(* IEC 61131-3 sources: LASAL/Network/HW_Network, 1 file *)

(* ---- ONE_HW_Network_Table.st ---- *)
#define OBJECTS_CONFIG

//Define part of class SdiasBase
//Address to access the Dataobject list via SPI SDO Read
#define SDIAS_SPI_DATA_OBJECT_LIST_PAGE_ADDRESS 16#FFFF
#define SDIAS_SPI_DATA_OBJECT_LIST_PAGE_OFFSET 16#00
#define SDIAS_SPI_DATA_OBJECT_LIST_IDENTIFIER 16#12345678

//Defines the number of optional list elements in the SPI List

#define SDIAS_SPI_NUMBER_OF_OPTIONAL_ELEMENTS 7

//#pragma message("EisMic 27.06.2014 14:44 \ Noch schauen ob ichs besser machen kann")
#define SDIAS_SPI_HEADER_BEFORE_OPTIONAL_ELEMENTS 16#18
#define SDIAS_SPI_HARDWARE_VERSION_OFFSET 16#C
#define SDIAS_SPI_VENDOR_ID_OFFSET 16#0

//SPI List IDs
#define SDIAS_SPI_IDENTIFICATION_LIST_ID 1
#define SDIAS_SPI_FLASH_CONFIGURATION_ID 2
#define SDIAS_SPI_VENDOR_NAME_ID 3
#define SDIAS_SPI_DEVICE_NAME_ID 4
#define SDIAS_SPI_SERIAL_NUMBER_ID 5
#define SDIAS_SPI_ORDERING_NUMBER_ID 6
#define SDIAS_SPI_DOCUMENTATION_PDF_ID 7
#define SDIAS_SPI_CALIB_DATA_ID 10
#define SDIAS_SPI_PDO_INFORMATION_ID 128
#include "..\..\Class\SdiasManager\SdiasManager.h"
#include "..\..\Class\SdiasBase\SdiasBase.h"
#include "..\..\Class\HwControl\HwControl.h"
#include "..\..\Source\interfaces\lsl_st_hardwaretree.h"
#include "..\..\Source\interfaces\lsl_st_mt.h"
//Define part of class _BusInterfaceSdiasDriveMng
#define BUSIF_SDIASDRIVEMNG_OFFSET_TYPELABEL        0x0000
#define BUSIF_SDIASDRIVEMNG_PARALIST_INDEX_SET      0x2210
#define BUSIF_SDIASDRIVEMNG_PARALIST_INDEX_INFO     0x2211
#define BUSIF_SDIASDRIVEMNG_PARALIST_INDEX_SETNR    174

#define BUSIF_SDIASDRIVEMNG_MAX_SERVICEBOX          4
#define BUSIF_SDIASDRIVEMNG_SDO_RESPONSE_TIMEOUT    SDIAS_SDO_TIMEOUT * 2
#define BUSIF_SDIASDRIVEMNG_SDO_TYPELABEL_TIMEOUT   10000  //10 sec timeout to read typelabel

#define BUSIF_SDIASDRIVEMNG_SDO_SERVICE_APP_MDD100        0x4150
#define BUSIF_SDIASDRIVEMNG_SDO_SERVICE_APP_LASAL         0x4C41
#define BUSIF_SDIASDRIVEMNG_SDO_SERVICE_APP_CANOPEN       0x4453
#define BUSIF_SDIASDRIVEMNG_SDO_SERVICE_APP_CANOPEN_LASAL 0x444C

#define BUSIF_SDIASDRIVEMNG_FULL_PARADATA_SIZE   12
#define BUSIF_SDIASDRIVEMNG_CANOPEN_FOOTER_SIZE   4
#define BUSIF_SDIASDRIVEMNG_LASAL_PARADATA_SIZE   4
#include "..\..\class\_drivemngbase\drivemngbase.h"
//Define part of class _DriveAxisBase
// Device ID for the Drive Cards
#define DRIVEMNG_AXISDEVICEID_SDD_OFFSET         0
#define DRIVEMNG_AXISEVICEID_MDD_OFFSET   16#10000
#define DRIVEMNG_AXISEVICEID_SDIAS_OFFSET 16#20000
#include "..\..\Class\_DriveMngBase\SDDDefinitions.h"
//Define part of class _DriveMngBase
#ifndef _T_DRIVEMNGBASE_H
#define _T_DRIVEMNGBASE_H

// DiasDrive Constants
#DEFINE SDDMAXENTRIES   32        // maximale Anzahl an Achsen
#DEFINE SDDMAXPLACE     3         // maximale Anzahl an Achsen pro Steckplatz

// Device ID for the Drive IF Cards
#define DRIVEMNG_BUSDEVICEID_VAC011    11
#define DRIVEMNG_BUSDEVICEID_VAC012  1061
#define DRIVEMNG_BUSDEVICEID_VAC013  1075

#define DRIVEMNG_BUSDEVICEID_MDD     1071

// Device ID for the Drive Cards
#define DRIVEMNG_DRVDEVICEID_SDD_OFFSET 0

#define DRIVEMNG_DRVDEVICEID_SDD305 DRIVEMNG_DRVDEVICEID_SDD_OFFSET + 16
#define DRIVEMNG_DRVDEVICEID_SDD310 DRIVEMNG_DRVDEVICEID_SDD_OFFSET +  3
#define DRIVEMNG_DRVDEVICEID_SDD315 DRIVEMNG_DRVDEVICEID_SDD_OFFSET +  1
#define DRIVEMNG_DRVDEVICEID_SDD335 DRIVEMNG_DRVDEVICEID_SDD_OFFSET + 12

#define DRIVEMNG_DRVDEVICEID_SDD205 DRIVEMNG_DRVDEVICEID_SDD_OFFSET + 22
#define DRIVEMNG_DRVDEVICEID_SDD210 DRIVEMNG_DRVDEVICEID_SDD_OFFSET +  9
#define DRIVEMNG_DRVDEVICEID_SDD215 DRIVEMNG_DRVDEVICEID_SDD_OFFSET +  5

#define DRIVEMNG_DRVDEVICEID_SDD105 DRIVEMNG_DRVDEVICEID_SDD_OFFSET + 21
#define DRIVEMNG_DRVDEVICEID_SDD115 DRIVEMNG_DRVDEVICEID_SDD_OFFSET + 10
#define DRIVEMNG_DRVDEVICEID_SDD120 DRIVEMNG_DRVDEVICEID_SDD_OFFSET +  7

#define DRIVEMNG_DRVDEVICEID_MDD_OFFSET 16#10000

#define DRIVEMNG_DRVDEVICEID_MDD111 DRIVEMNG_DRVDEVICEID_MDD_OFFSET + 1
#define DRIVEMNG_DRVDEVICEID_MDD121 DRIVEMNG_DRVDEVICEID_MDD_OFFSET + 2

#define DRIVEMNG_DRVDEVICEID_SDIAS_OFFSET 16#20000

#define DRIVEMNG_DRVDEVICEID_DC061 DRIVEMNG_DRVDEVICEID_SDIAS_OFFSET + 16#180 // 1 = 1 Achse 80 SDIAS

#define DRIVEMNG_DRIVESCOPE_GETALL_PARAM    16#2080
#define DRIVEMNG_DRIVESCOPE_SCOPE_BIT       16#60000000
#define DRIVEMNG_DRIVESCOPE_SINDEX_RANGE    511

#endif // _T_DRIVEMNGBASE_H
//Define part of class BusInterfaceSDIASInternal
#define BUSIF_INTERNAL_MAX_NR_DO 100

// Defines for Mutex Generation
#define INTERNAL_STR_MUTEX_NAME_SEPERATOR ".."
#define INTERNAL_MUTEX_NAME_END_LENGTH 5
#define INTERNAL_MUTEX_NAME_MAX_LENGTH 32
#include "..\..\Source\BusInterface.h"
//Define part of class DM161
#define DEVICE_ID_DM161 1029
#include "..\..\Class\HwControl\watchdog.h"
#include "..\..\Source\interfaces\lsl_st_sysinfo.h"
#include "..\..\Source\interfaces\lsl_st_systrace.h"
#include <.\lsl_st_mt.h>
//Define part of class SafetyUDP
#define SAFETY_UDP_MAX_SOCKETS                6     // Max number of socket

#define SAFETY_UDP_CLT_SEND_OK                0    // Send ok
#define SAFETY_UDP_CLT_INVALID_HANDLE        -1    // Invalid handle
#define SAFETY_UDP_CLT_NOT_OPEN              -2    // Socket is not open
#define SAFETY_UDP_CLT_SEND_FAILED           -3    // Send failed
#define SAFETY_UDP_CLT_SEND_BUFFER_FULL      -4    // Send buffer is full
#define SAFETY_UDP_CLT_DATA_TO_BIG           -5    // Data to big

#define SAFETY_UDP_MAXIMUM_SEGMENT_SIZE    1452    // Maximum of user data

#define SAFETY_UDP_TIMEOUT_OPENSOCKET    (1000)    //timeout for opening socket

#define SAFETY_UDP_RECEIVE_TIMEOUT          800

#define SAFETY_UDP_TX_BUFFER_SIZE          1024
//Define part of class SafetyManager
#define LogBufferSize 1000
#include "..\..\Class\SafetyManager\SafetyManager.h"
#include "..\..\Source\interfaces\lsl_st_safetydll.h"
//Define part of class SdiasManager
#define SDIAS_SDO_MAX_LENGTH              128
#define SDIAS_SDO_RINGBUFFER_NO            64
#define SDIAS_SDO_CHANNEL_NO                3   // fixed in the VI hardware to be 3

// watchdog trigger interval (after 130ms of no trigger the SDIAS HW goes into reset again and takes at least another 10ms to be ready again)
#define SDIAS_WATCHDOG_TRIGGER_TIME        40

// time needed by sdias modules to start up after the watchdog is triggered the first time in ms
#define SDIAS_HARDWARE_STARTUP_TIME        15

// sdias manager needs 2 ticks to handle event for read task (measure sync time)
#define SDIAS_SYNC_MEASURE_TICKS            2

// after activating the PLL SyncOut it takes 3 cycles until the SDIAS sync can be injected
#define SDIAS_CYCLES_WAIT_AFTER_SYNC_ENABLE 3

// wait 1 bus cycle at start to get valid numbers in the task info
#define SDIAS_TASKINFO_READY_TICKS          1

// time to wait (in ms) until other tasks in the same or lower priority than post init have done their stuff
#define SDIAS_WAIT_TIME_IN_POST_INIT        1

#define SIZE_PER_SDIAS_CLIENT               16#0400

// for far memory accesses: 1 module can hold maximum 256 1K blocks (0-255)
#define SDIAS_1K_BLOCK_NO                       256

// far memory accesses maximum length in bytes
#define SDIAS_MAX_SIZE_FAR_MEM_ACCESS           127

#define SDIAS_OFFSET_HW_CONFIG              16#FF00
#define SDIAS_OFFSET_TASK_EVENT_IDS         16#FF10
#define SDIAS_OFFSET_FEATURE_INFO           16#FF18
#define SDIAS_OFFSET_APPLI_LED_STATES       16#FF20
#define SDIAS_OFFSET_SYNC_INJECTION_CFG     16#FF3D
#define SDIAS_OFFSET_TRIGGER_UNIT_SETUP_0   16#FF41
#define SDIAS_OFFSET_TRIGGER_UNIT_SETUP_1   16#FF45
#define SDIAS_OFFSET_TASK_START_CFG_0       16#FF60
#define SDIAS_OFFSET_TASK_CONFIG_0          16#FF86
#define SDIAS_OFFSET_TASK_CONFIG_1          16#FF96
#define SDIAS_OFFSET_TASK_INFO_1            16#FF94
#define SDIAS_OFFSET_TASK_HANDSHAKE_1       16#FF9B
#define SDIAS_OFFSET_TASK_DURATION_TIME_1   16#FF9C
#define SDIAS_OFFSET_TASK_DURATION_TIME_2   16#FFAC
#define SDIAS_OFFSET_TASK_CONFIG_2          16#FFA6

#define SDIAS_RETRIES_ALLOWED         2

// mask to get global error flag out of message counter byte of SDO responses
#define SDIAS_MASK_GLOBAL_ERROR_FLAG        16#80

// mask to get message counter out of message counter byte of SDO responses
#define SDIAS_MASK_MESSAGE_COUNTER          16#3F

#define SDIAS_EVENT_MASK_ID_SYNC_OUT0       16#10
#define SDIAS_EVENT_MASK_ID_SYNC_OUT1       16#11
#define SDIAS_EVENT_MASK_ID_SYNC_OUT2       16#12
#define SDIAS_EVENT_MASK_ID_SYNC_OUT3       16#13

#define SDIAS_MANAGER_SYNC_SYNCOUT_ID       16#85
#define SDIAS_TASK_START_EVENT_SYNCOUT_ID   16#86

#define SDIAS_PLACE_NO_MODULE_ADDED_SO_FAR  16#80000000

#define SDIAS_TRIGGER_UNIT_BYTE_SIZE        2

#define SDIAS_WAIT_TIME_FIRMWARE_HANDSHAKE  5 * 1000

// if the firmware version is below this, there might be problems with SCP111 and other modules => print warning at startup
#define SDIAS_FW_VERSION_SDO_ERROR_FIXED    16#120

// if the protocol version ist below this, Control Read/Broadcast Write Command is not supported by sdiasmanager
#define SDIAS_PROTOCOLVERSION_BROADCAST     16#120

// if the cil version ist below this, Control Read/Broadcast Write Command is not supported by OS for local SDIAS.
#define SDIAS_CILVERSION_BROADCAST         16#5001

// timeout for blocking the init during initialisation (in ms)
#define SDIAS_INIT_BLOCK_TIMEOUT            20 * 1000

#define SDIAS_MUTEX_NAME_END_LENGTH 3
#define SDIAS_MUTEX_NAME_MAX_LENGTH 32
#define SDIAS_MUTEX_STR_SEPERATOR   ".."

//#define SDIAS_RT_TIME_MEASUREMENT
#ifdef SDIAS_RT_TIME_MEASUREMENT
  #pragma message("ATTENTION: SDIAS real time measurement is active and needs additional ressources in the realtime task")
#endif

(* SDIAS data object commands  *)
#define	 SDIAS_CMD_END							  0x00			(* End command										          *)
#define	 SDIAS_CMD_ACC_MEMORY				  0x01			(* Access dpram memory								      *)
#define	 SDIAS_CMD_ACC_CONTROL				0x02			(* Access dpram control memory						  *)
#define	 SDIAS_CMD_GLOBAL						  0x03			(* SDIAS global command								      *)
#define	 SDIAS_CMD_COPY_LOCAL					0x04			(* DPRAM copy command in local dpram				*)
#define	 SDIAS_CMD_JMP_LOCAL					0x05			(* DPRAM jump command in local dpram 				*)
#define  SDIAS_CMD_ACC_MEMORY_FAR     0x07      (* SDIAS Far Memory Access                  *)

(* SDIAS defines for data object handling *)
// Write data oject list
#define	 SDIAS_DOL_WRITE_USAGE_DOL_EMPTY	  0x20			(* Usage of empty write dol list (wachtdog trigger + end command)   *)
#define	 SDIAS_DOL_WRITE_USAGE_DTA_EMPTY	  0x03			(* Usage of empty write dol data (DO ctrl of 2x copy command for task information + DO ctrl of watchdog trigger      *)
#define	 SDIAS_DOL_WRITE_OFFSET_END_CMD			0x10			(* One data object in list - offset = 1 DO size = 0x10						  *)
#define	 SDIAS_DOL_WRITE_OFFSET_FIRST_DTA		0x02			(* Offset of first data byte of second copy command = 2 (DO ctrl)   *)
#define	 SDIAS_DOL_WRITE_OFFSET_LAST_DTA		0x02			(* Offset of last data byte of second copy command = 2 (DO ctrl )   *)

// Read data oject list
#define	 SDIAS_DOL_READ_USAGE_DOL_EMPTY	    0x30			(* Usage of empty read dol list (2x task info copy command + end command)   *)
#define	 SDIAS_DOL_READ_USAGE_DTA_EMPTY	    0x0D			(* Usage of empty write dol data (DO ctrl of 2x copy command for task information + DO ctrl of watchdog trigger      *)
#define	 SDIAS_DOL_READ_OFFSET_END_CMD			0x20			(* One data object in list - offset = 1 DO size = 0x10						          *)
#define	 SDIAS_DOL_READ_OFFSET_FIRST_DTA		0x07			(* Offset of first data byte of second copy command = 7 = DO state          *)
#define	 SDIAS_DOL_READ_OFFSET_LAST_DTA		  0x0C			(* Offset of last data byte of second copy command = 12 (last byte of task information)       *)

//Versionsnumber where SDIAS SPI Read Accesses are available
#define  SDIAS_SDO_SPI_FIRMWARE_VERSION_AVAILABLE 16#0120

//error info mask
#define  SDIAS_ERROR_INFO_MASK    2#1000011000011111

// Broadcast DO Info
#define SDIAS_OFFSET_CLIENT_CTRLTIMESTAMP   16#0190
#define SDIAS_NR_TIMEBROADCAST_DOS 2
#define SDIAS_TIMEBROADCAST_SUBCMD 16#B0
#include "..\..\Source\interfaces\lsl_st_pll.h"
//Define part of class SdiasPLC
#define SDIASM_OBJECT_PATH            16#88000002   // Object Path for VSDIASmanager Length = 2 (First 2byte), Domain = 0 (3rd byte), Escape Sequence SDIAS (4th byte)
//Define part of class SR022
#define DEVICE_ID_SR022             1083        //DeviceID of SR022

#define SR022_ADDR_CYC_WRITE        16#00       //Address for TPDO
#define SR022_ADDR_CYC_READ         16#08       //Address for RPDO

#define SR022_ADDR_CFG_FIRMWARE     16#200      //Address-Offset to the Configuration of the Firmware
#define SR022_ADDR_STATE_FIRMWARE   16#280      //Address-Offset to the Status of the Firmware
#define SR022_ADDR_READ_SDO         16#0C       //Address-Offset read sdo data
#define SR022_ADDR_I2T_THRESHOLD    16#18       //Address-Offset to I²T Threshold
#define SR022_ADDR_DC_SEQUENCER     16#20       //Address-Offset to sequencer SR022

#define SR022_INVALID_VALUE         16#80000010$DINT

#define SR022_NOENCODER             0
#define SR022_TTL_MODE              1
#define SR022_RS422_MODE            2

//Define for the H-Bridge
//-----------------------------------------------------------
#define SR022_GATE_A_LOW		          2#0100000000000000    //Bit-Configuration for Enable GateA Low-Switch
#define SR022_GATE_A_HIGH		          2#0001000000000000    //Bit-Configuration for Enable GateA High-Switch
#define SR022_GATE_B_LOW		          2#1000000000000000    //Bit-Configuration for Enable GateB Low-Switch
#define SR022_GATE_B_HIGH		          2#0010000000000000    //Bit-Configuration for Enable GateB High-Switch

#define SR022_MASK_CONTROL	          16#0FFF     //Mask for Output Sequence Bits
#define SR022_MASK_TIME		            16#F000     //Mask for TimeValue

#define SR022_T_SWITCH                41      //Delay Time for Switch
#define SR022_DEFAULT_SEQ_INIT        1       //Initilization for Sequencer => After 1 FPGA-Cycle switch to next Sequency

#define SR022_FPGA_FREQ_MHZ           50    //Frequency of FPGA

#define SR022_SDO_RESPONSE_TIMEOUT  SDIAS_SDO_TIMEOUT * 2     //SDO-Response Timeout

//#define SR022_I2T_THRESHOLD          16000000   //Maximal allowed I²T Value in mA²s ==> 16 A²s
//#pragma message ("TarPet: dieser Wert wurde vorest empirisch ermittelt und sollte noch genau bestimmt werden");
#define SR022_I2T_THRESHOLD          78000   //Maximal allowed I²T Value in mA²s ==> 16 A²s

#define SR022_SPEED_SCALING          10000      //Scaling of the Server Speed (0.00% to 100.00%)
#define SR022_MINPULSE_SCALING       1000       //Scaling of the Server MinPulse (0.0% to 100.0%)
//Define part of class ST011
#define DEVICE_ID_ST011 1052
#define ST011_MINIMAL_PULSEWIDTH 16#003C

#define ST011_ADDR_PDO_WRITE    16#001F
#define ST011_ADDR_SDO_WRITE_1  16#0025
#define ST011_ADDR_PDO_READ     16#0037
#define ST011_ADDR_SDO_WRITE_2  16#0042

#define ST011_FPGAVersion_PulsCntCorrect 16#12

// in MHz
#define ST011_FREQUENCY_MHZ 125

// in Hz
#define ST011_FREQUENCY_HZ (ST011_FREQUENCY_MHZ * 1000000)

#define ST011_SDO_RESPONSE_TIMEOUT  SDIAS_SDO_TIMEOUT * 2
//Define part of class ST151Base
#define DEVICE_ID_ST151                                                    1086

#define ST151_ADDR_PDO_WRITE                                            16#0000
#define ST151_ADDR_PDO_READ                                             16#0038
#define ST151_ADDR_SDO_1                                                16#0008
#define ST151_ADDR_SDO_2           (ST151_ADDR_SDO_1+sizeof(t_s_ConfigModule1))
#define ST151_ADDR_SDO_3                                (ST151_ADDR_PDO_READ+6)  //only read sdo!!!
#define ST151_ADDR_SDO_4           (ST151_ADDR_SDO_3+sizeof(t_s_ConfigModule3))
#define ST151_ADDR_SDO_5           (ST151_ADDR_SDO_4+sizeof(t_s_ConfigModule4))
#define ST151_ADDR_SDO_6           (ST151_ADDR_SDO_5+sizeof(t_s_ConfigModule5))

#define ST151_OSZI_ADDR_WRITE                                           16#0800
#define ST151_OSZI_ADDR_READ                                            16#0808
#define ST151_OSZI_ADDR_DATA                                            16#0820
#define ST151_OSZI_READPOINTER_OFFSET                                   16#0020
#define ST151_OSZI_ONE_PDOSIZE                                              126
#define ST151_OSZI_VALUES_DATA             (ST151_OSZI_ONE_PDOSIZE/sizeof(UINT))
#define ST151_OSZI_BUFFER_SIZE                                             1024
#define ST151_OSZI_MAX_SAMPLES             (ST151_OSZI_BUFFER_SIZE/sizeof(UINT))
#define ST151_OSZI_MAX_PDOREAD   ((ST151_OSZI_BUFFER_SIZE/ST151_OSZI_ONE_PDOSIZE)+1)

// in MHz
#define ST151_FREQUENCY_MHZ                             125
// in Hz
#define ST151_FREQUENCY_HZ   (ST151_FREQUENCY_MHZ * 1000000)

#define ST151_SDO_RESPONSE_TIMEOUT   (SDIAS_SDO_TIMEOUT * 2)
#define ST151_SDO_MAX_RETRYS                              3

#define ST151_MAXFREQUENCY_OUT                   2_000_000 // 2Mhz/64 max frequency of module output
#define ST151_MAXSTEPPING_MODES                          6
#define ST151_FREQLIMITS_TABLESIZE      (ST151_MAXSTEPPING_MODES*sizeof(UDINT)*2)

#define ST151_MAX_ALLOWED_PERCENT                      100 // maximum value for percent value
#define ST151_BLANKING_TIME                             10 // minimum on time of pwm (*20ns)

#define ST151_CYCLICREFRESHDATA_TIME                   200 // time to refresh asynchrone values
#define ST151_INVALID_VALUE                   16#8000_0010 // invalid value for server
#define ST151_AUTOSET_FREQUENCYLIMIT          16#0000_0000 // value for autoset limit
#define ST151_DEACTIVATE_FREQUENCYLIMIT       16#FFFF_FFFF // value for deactivate limit

#define ST151_MAX_ALLOWED_CURRENT                     5000 // max allowed current (5A) in mA, from h-bridge according to hw-documentation
#define ST151_MAX_ALLOWED_CHOPPEROFFTIME              2500 // max allowed chopper off time in 20ns steps
#define ST151_MIN_ALLOWED_CHOPPEROFFTIME              1500 // min allowed chopper off time in 20ns steps
#define ST151_STALL_CURRENT_LIMIT                     1000 // calculation for stall current in permille
#define ST151_CURRENTOFFSETADJUST_MAX                  250 // maximum current offset adjust in mA
#define ST151_CURRENTOFFSETADJUST_MIN                 -250 // minimum current offset adjust in mA

//pll settings
#define ST151_SYNC_OUT_ID                             16#03
#define ST151_PLL_OFFSET                             16#140
#define ST151_PLL_CONTROL               (ST151_PLL_OFFSET+8)

#define ST151_ERROR_BITMASK_STATE_WORD               0x013E
#define ST151_ERROR_BITMASK_EXTENDED_STATE_WORD      0xFF3E
//Define part of class VaranManager
#define SIZE_PAYLOAD_FRAME_HEADER_DO      16#38  // Const because datasize is in the Payload DOs
#define SIZE_PAYLOAD_IRQ_FRAME_HEADER_DO  16#40  // Const because datasize is in the Payload DOs

#define VM_MAX_POST_INIT_MODULES  1000

#define VM_OBJECT_PATH            16#81000002   // Object Path for Varanmanager Length = 2 (First 2byte), Domain = 0 (3rd byte), Escape Sequence Varan (4th byte)
#include "..\..\Class\VaranManager\VaranManager.h"
#include "..\..\Source\interfaces\lsl_st_kernel.h"

FUNCTION GLOBAL TAB ONE_HW_Network
-1$UINT, 0$UINT,
0$UINT, 0$UINT,

39$UDINT,
TO_UDINT(1048633017), "_BusInterfaceSdiasDriveMng", 1$UINT, 10$UINT, 4$UINT,
TO_UDINT(529317953), "_CanLib", 1$UINT, 10$UINT, 2$UINT,
TO_UDINT(912370472), "_DriveAxis", 1$UINT, 63$UINT, 4$UINT,
TO_UDINT(4124502522), "_DriveAxisBase", 1$UINT, 72$UINT, 0$UINT,
TO_UDINT(833307860), "_DriveAxisSet", 1$UINT, 20$UINT, 4$UINT,
TO_UDINT(1470062879), "_DriveMng_DC062", 1$UINT, 16$UINT, 4$UINT,
TO_UDINT(496739206), "_DriveMngBase", 1$UINT, 41$UINT, 0$UINT,
TO_UDINT(4078275645), "_SerLib", 1$UINT, 34$UINT, 2$UINT,
TO_UDINT(2897291062), "ASCII_BIN", 1$UINT, 21$UINT, 1$UINT,
TO_UDINT(3882880897), "BusInterfaceSDIASInternal", 2$UINT, 0$UINT, 0$UINT,
TO_UDINT(658879389), "CP112_IOs", 1$UINT, 0$UINT, 1$UINT,
TO_UDINT(794617671), "CriticalSection", 0$UINT, 4$UINT, 2$UINT,
TO_UDINT(4282685340), "DM161", 1$UINT, 12$UINT, 1$UINT,
TO_UDINT(3238133653), "Hub_Base", 1$UINT, 21$UINT, 0$UINT,
TO_UDINT(1770276445), "Hub_Base_Root", 2$UINT, 11$UINT, 1$UINT,
TO_UDINT(2471641665), "HwControl", 5$UINT, 2$UINT, 1$UINT,
TO_UDINT(1193052171), "HwControlBase", 1$UINT, 10$UINT, 0$UINT,
TO_UDINT(4260294091), "HWRtPostScan", 1$UINT, 0$UINT, 1$UINT,
TO_UDINT(2225119864), "MerkerEx", 1$UINT, 22$UINT, 21$UINT,
TO_UDINT(933570811), "RAMex", 1$UINT, 17$UINT, 4$UINT,
TO_UDINT(1799751072), "SafetyManager", 2$UINT, 11$UINT, 1$UINT,
TO_UDINT(3727715967), "SafetyUDP", 1$UINT, 2$UINT, 0$UINT,
TO_UDINT(3175101883), "SdiasBase", 1$UINT, 58$UINT, 0$UINT,
TO_UDINT(4173303375), "SdiasHubBase", 1$UINT, 10$UINT, 1$UINT,
TO_UDINT(2118381352), "SdiasManager", 1$UINT, 92$UINT, 1$UINT,
TO_UDINT(1159122596), "SdiasPLC", 2$UINT, 0$UINT, 1$UINT,
TO_UDINT(2317024038), "SetCurrent", 0$UINT, 0$UINT, 1$UINT,
TO_UDINT(3646514510), "SR022", 1$UINT, 2$UINT, 1$UINT,
TO_UDINT(1310079211), "ST011", 1$UINT, 11$UINT, 1$UINT,
TO_UDINT(733517784), "ST151", 1$UINT, 2$UINT, 2$UINT,
TO_UDINT(1691609973), "ST151_IntVisu", 1$UINT, 0$UINT, 2$UINT,
TO_UDINT(1832775974), "ST151Base", 1$UINT, 2$UINT, 0$UINT,
TO_UDINT(1850111279), "String", 1$UINT, 10$UINT, 17$UINT,
TO_UDINT(2898603620), "StringInternal", 1$UINT, 82$UINT, 0$UINT,
TO_UDINT(2940693151), "VaranManager", 3$UINT, 1$UINT, 0$UINT,
TO_UDINT(1989862026), "VaranManager_1", 2$UINT, 1$UINT, 1$UINT,
TO_UDINT(4035182347), "VaranManager_Base", 1$UINT, 24$UINT, 0$UINT,
TO_UDINT(3232495061), "VirtualBaseInit", 1$UINT, 3$UINT, 0$UINT,
TO_UDINT(819479645), "XXXBase_IOs", 1$UINT, 0$UINT, 0$UINT,

1$UINT, TO_UDINT(1755887647), "_DRIVEMNG_DC0621\BUSINTERFACESDIASDRIVEMNG",
1$UINT, TO_UDINT(3678180828), "_DRIVEMNG_DC0622\BUSINTERFACESDIASDRIVEMNG",
1$UINT, TO_UDINT(3048246941), "_DRIVEMNG_DC0623\BUSINTERFACESDIASDRIVEMNG",
1$UINT, TO_UDINT(1734723611), "_DRIVEMNG_DC0624\BUSINTERFACESDIASDRIVEMNG",

1$UINT, TO_UDINT(3194356815), "CP112_IOS1\_BASE\_CANLIB1",
1$UINT, TO_UDINT(661607925), "CP112_IOS1\_BASE\_CANLIB2",

_NO_ATTR, TO_UDINT(3059689190), "_DRIVEAXIS1",
_NO_ATTR, TO_UDINT(794195804), "_DRIVEAXIS2",
_NO_ATTR, TO_UDINT(1481721802), "_DRIVEAXIS3",
_NO_ATTR, TO_UDINT(3325416041), "_DRIVEAXIS4",

1$UINT, TO_UDINT(4275951967), "_DRIVEAXIS1\SDDAXSET1",
1$UINT, TO_UDINT(1732231006), "_DRIVEAXIS2\SDDAXSET1",
1$UINT, TO_UDINT(2796642462), "_DRIVEAXIS3\SDDAXSET1",
1$UINT, TO_UDINT(2408215837), "_DRIVEAXIS4\SDDAXSET1",

_NO_ATTR, TO_UDINT(243498275), "_DRIVEMNG_DC0621",
_NO_ATTR, TO_UDINT(2542415001), "_DRIVEMNG_DC0622",
_NO_ATTR, TO_UDINT(3767344143), "_DRIVEMNG_DC0623",
_NO_ATTR, TO_UDINT(2129234348), "_DRIVEMNG_DC0624",

1$UINT, TO_UDINT(3879313428), "CP112_IOS1\_BASE\_SERLIB1",
1$UINT, TO_UDINT(2117136814), "CP112_IOS1\_BASE\_SERLIB2",

1$UINT, TO_UDINT(3603645853), "VARANMANAGER_11\_BASE\ASCII_BIN1",

_NO_ATTR, TO_UDINT(222643709), "CP112_IOS1",

1$UINT, TO_UDINT(2972590922), "HWCONTROL1\SAFETYMANAGER\UDPRECEIVEDATA",
1$UINT, TO_UDINT(1868223583), "HWCONTROL1\SAFETYMANAGER\UDPSENDDATA",

_NO_ATTR, TO_UDINT(2056942671), "DM1611",

1$UINT, TO_UDINT(1776428101), "VARANMANAGER_11\HUB_BASE_ROOT0",

_NO_ATTR, TO_UDINT(2190789875), "HWCONTROL1",

1$UINT, TO_UDINT(1673205898), "HWCONTROL1\HWRTPOSTSCAN",

1$UINT, TO_UDINT(1089285877), "DM1611\_BASE\SERIALNOSTR\MERKEREX0",
1$UINT, TO_UDINT(566457232), "SR0221\_BASE\SERIALNOSTR\MERKEREX0",
1$UINT, TO_UDINT(3227848145), "ST0111\_BASE\SERIALNOSTR\MERKEREX0",
1$UINT, TO_UDINT(921637672), "ST1511\_BASE\_BASE\SERIALNOSTR\MERKEREX0",
1$UINT, TO_UDINT(3174837553), "ST1512\_BASE\_BASE\SERIALNOSTR\MERKEREX0",
1$UINT, TO_UDINT(3868254288), "_DRIVEAXIS1\MERKEREX2",
1$UINT, TO_UDINT(2138211921), "_DRIVEAXIS2\MERKEREX2",
1$UINT, TO_UDINT(3204209041), "_DRIVEAXIS3\MERKEREX2",
1$UINT, TO_UDINT(2546420754), "_DRIVEAXIS4\MERKEREX2",
1$UINT, TO_UDINT(1361534785), "_DRIVEMNG_DC0621\BUSINTERFACESDIASDRIVEMNG\_BASE\SERIALNOSTR\MERKEREX0",
1$UINT, TO_UDINT(570430050), "_DRIVEMNG_DC0621\FWDATESTRING\MERKEREX0",
1$UINT, TO_UDINT(1339808896), "_DRIVEMNG_DC0621\FWNUMSTRING\MERKEREX0",
1$UINT, TO_UDINT(925076081), "_DRIVEMNG_DC0622\BUSINTERFACESDIASDRIVEMNG\_BASE\SERIALNOSTR\MERKEREX0",
1$UINT, TO_UDINT(2048834378), "_DRIVEMNG_DC0622\FWDATESTRING\MERKEREX0",
1$UINT, TO_UDINT(960423357), "_DRIVEMNG_DC0622\FWNUMSTRING\MERKEREX0",
1$UINT, TO_UDINT(354433377), "_DRIVEMNG_DC0623\BUSINTERFACESDIASDRIVEMNG\_BASE\SERIALNOSTR\MERKEREX0",
1$UINT, TO_UDINT(4215004781), "_DRIVEMNG_DC0623\FWDATESTRING\MERKEREX0",
1$UINT, TO_UDINT(2722959209), "_DRIVEMNG_DC0623\FWNUMSTRING\MERKEREX0",
1$UINT, TO_UDINT(4213841937), "_DRIVEMNG_DC0624\BUSINTERFACESDIASDRIVEMNG\_BASE\SERIALNOSTR\MERKEREX0",
1$UINT, TO_UDINT(3391351066), "_DRIVEMNG_DC0624\FWDATESTRING\MERKEREX0",
1$UINT, TO_UDINT(3572799431), "_DRIVEMNG_DC0624\FWNUMSTRING\MERKEREX0",

1$UINT, TO_UDINT(3414815221), "_DRIVEAXIS1\RAMEX2",
1$UINT, TO_UDINT(1158084118), "_DRIVEAXIS2\RAMEX2",
1$UINT, TO_UDINT(2309813896), "_DRIVEAXIS3\RAMEX2",
1$UINT, TO_UDINT(2204762001), "_DRIVEAXIS4\RAMEX2",

1$UINT, TO_UDINT(1778590035), "HWCONTROL1\SAFETYMANAGER",

1$UINT, TO_UDINT(1007630054), "SDIASPLC1\SDIASHUBBASE1",

1$UINT, TO_UDINT(4015996540), "SDIASPLC1\SDIASMANAGER1",

_NO_ATTR, TO_UDINT(1378000520), "SDIASPLC1",

_NO_ATTR, TO_UDINT(1364947121), "SETCURRENT1",

_NO_ATTR, TO_UDINT(308402757), "SR0221",

_NO_ATTR, TO_UDINT(3024798335), "ST0111",

_NO_ATTR, TO_UDINT(201264582), "ST1511",
_NO_ATTR, TO_UDINT(2465619068), "ST1512",

1$UINT, TO_UDINT(869501406), "ST1511\ST151_INTVISU1",
1$UINT, TO_UDINT(437992748), "ST1512\ST151_INTVISU1",

1$UINT, TO_UDINT(2011818843), "DM1611\_BASE\SERIALNOSTR",
1$UINT, TO_UDINT(3834696548), "SR0221\_BASE\SERIALNOSTR",
1$UINT, TO_UDINT(3723324983), "ST0111\_BASE\SERIALNOSTR",
1$UINT, TO_UDINT(3070230801), "ST1511\_BASE\_BASE\SERIALNOSTR",
1$UINT, TO_UDINT(2196617026), "ST1512\_BASE\_BASE\SERIALNOSTR",
1$UINT, TO_UDINT(189353776), "_DRIVEMNG_DC0621\BUSINTERFACESDIASDRIVEMNG\_BASE\SERIALNOSTR",
1$UINT, TO_UDINT(275191107), "_DRIVEMNG_DC0621\FWDATESTRING",
1$UINT, TO_UDINT(1236665617), "_DRIVEMNG_DC0621\FWNUMSTRING",
1$UINT, TO_UDINT(880947621), "_DRIVEMNG_DC0622\BUSINTERFACESDIASDRIVEMNG\_BASE\SERIALNOSTR",
1$UINT, TO_UDINT(1812344984), "_DRIVEMNG_DC0622\FWDATESTRING",
1$UINT, TO_UDINT(4101794271), "_DRIVEMNG_DC0622\FWNUMSTRING",
1$UINT, TO_UDINT(2534676969), "_DRIVEMNG_DC0623\BUSINTERFACESDIASDRIVEMNG\_BASE\SERIALNOSTR",
1$UINT, TO_UDINT(4043952622), "_DRIVEMNG_DC0623\FWDATESTRING",
1$UINT, TO_UDINT(703246426), "_DRIVEMNG_DC0623\FWNUMSTRING",
1$UINT, TO_UDINT(1259654287), "_DRIVEMNG_DC0624\BUSINTERFACESDIASDRIVEMNG\_BASE\SERIALNOSTR",
1$UINT, TO_UDINT(2495904558), "_DRIVEMNG_DC0624\FWDATESTRING",
1$UINT, TO_UDINT(1419359746), "_DRIVEMNG_DC0624\FWNUMSTRING",

_NO_ATTR, TO_UDINT(2395414379), "VARANMANAGER_11",

//Internal connections
0$UDINT,
64$UDINT,
TO_UDINT(0), "SerialNoStr", TO_UDINT(69),
TO_UDINT(1), "SerialNoStr", TO_UDINT(72),
TO_UDINT(2), "SerialNoStr", TO_UDINT(75),
TO_UDINT(3), "SerialNoStr", TO_UDINT(78),
TO_UDINT(6), "SDDAxSet1", TO_UDINT(10),
TO_UDINT(6), "MerkerEx2", TO_UDINT(33),
TO_UDINT(6), "RAMex2", TO_UDINT(49),
TO_UDINT(7), "SDDAxSet1", TO_UDINT(11),
TO_UDINT(7), "MerkerEx2", TO_UDINT(34),
TO_UDINT(7), "RAMex2", TO_UDINT(50),
TO_UDINT(8), "SDDAxSet1", TO_UDINT(12),
TO_UDINT(8), "MerkerEx2", TO_UDINT(35),
TO_UDINT(8), "RAMex2", TO_UDINT(51),
TO_UDINT(9), "SDDAxSet1", TO_UDINT(13),
TO_UDINT(9), "MerkerEx2", TO_UDINT(36),
TO_UDINT(9), "RAMex2", TO_UDINT(52),
TO_UDINT(14), "FWDateString", TO_UDINT(70),
TO_UDINT(14), "FWNumSTring", TO_UDINT(71),
TO_UDINT(14), "BusInterfaceSdiasDriveMng", TO_UDINT(0),
TO_UDINT(15), "FWDateString", TO_UDINT(73),
TO_UDINT(15), "FWNumSTring", TO_UDINT(74),
TO_UDINT(15), "BusInterfaceSdiasDriveMng", TO_UDINT(1),
TO_UDINT(16), "FWDateString", TO_UDINT(76),
TO_UDINT(16), "FWNumSTring", TO_UDINT(77),
TO_UDINT(16), "BusInterfaceSdiasDriveMng", TO_UDINT(2),
TO_UDINT(17), "FWDateString", TO_UDINT(79),
TO_UDINT(17), "FWNumSTring", TO_UDINT(80),
TO_UDINT(17), "BusInterfaceSdiasDriveMng", TO_UDINT(3),
TO_UDINT(21), "_SerLib1", TO_UDINT(18),
TO_UDINT(21), "_SerLib2", TO_UDINT(19),
TO_UDINT(21), "_CanLib1", TO_UDINT(4),
TO_UDINT(21), "_CanLib2", TO_UDINT(5),
TO_UDINT(24), "SerialNoStr", TO_UDINT(64),
TO_UDINT(26), "SafetyManager", TO_UDINT(53),
TO_UDINT(26), "HWRtPostScan", TO_UDINT(27),
TO_UDINT(53), "UdpSendData", TO_UDINT(23),
TO_UDINT(53), "UdpReceiveData", TO_UDINT(22),
TO_UDINT(56), "SdiasManager1", TO_UDINT(55),
TO_UDINT(56), "SdiasHubBase1", TO_UDINT(54),
TO_UDINT(58), "SerialNoStr", TO_UDINT(65),
TO_UDINT(59), "SerialNoStr", TO_UDINT(66),
TO_UDINT(60), "SerialNoStr", TO_UDINT(67),
TO_UDINT(60), "ST151_IntVisu1", TO_UDINT(62),
TO_UDINT(61), "SerialNoStr", TO_UDINT(68),
TO_UDINT(61), "ST151_IntVisu1", TO_UDINT(63),
TO_UDINT(64), "MerkerEx0", TO_UDINT(28),
TO_UDINT(65), "MerkerEx0", TO_UDINT(29),
TO_UDINT(66), "MerkerEx0", TO_UDINT(30),
TO_UDINT(67), "MerkerEx0", TO_UDINT(31),
TO_UDINT(68), "MerkerEx0", TO_UDINT(32),
TO_UDINT(69), "MerkerEx0", TO_UDINT(37),
TO_UDINT(70), "MerkerEx0", TO_UDINT(38),
TO_UDINT(71), "MerkerEx0", TO_UDINT(39),
TO_UDINT(72), "MerkerEx0", TO_UDINT(40),
TO_UDINT(73), "MerkerEx0", TO_UDINT(41),
TO_UDINT(74), "MerkerEx0", TO_UDINT(42),
TO_UDINT(75), "MerkerEx0", TO_UDINT(43),
TO_UDINT(76), "MerkerEx0", TO_UDINT(44),
TO_UDINT(77), "MerkerEx0", TO_UDINT(45),
TO_UDINT(78), "MerkerEx0", TO_UDINT(46),
TO_UDINT(79), "MerkerEx0", TO_UDINT(47),
TO_UDINT(80), "MerkerEx0", TO_UDINT(48),
TO_UDINT(81), "ASCII_BIN1", TO_UDINT(20),
TO_UDINT(81), "Hub_Base_Root0", TO_UDINT(25),
0$UDINT,
69$UDINT,
TO_UDINT(6), "DriveMng", TO_UDINT(14), "CmdState",
TO_UDINT(6), "DriveAxisSet", TO_UDINT(10), "Server0",
TO_UDINT(7), "DriveMng", TO_UDINT(15), "CmdState",
TO_UDINT(7), "DriveAxisSet", TO_UDINT(11), "Server0",
TO_UDINT(8), "DriveMng", TO_UDINT(16), "CmdState",
TO_UDINT(8), "DriveAxisSet", TO_UDINT(12), "Server0",
TO_UDINT(9), "DriveMng", TO_UDINT(17), "CmdState",
TO_UDINT(9), "DriveAxisSet", TO_UDINT(13), "Server0",
TO_UDINT(10), "coMerkerEx", TO_UDINT(33), "m_udLength",
TO_UDINT(10), "coRamEx", TO_UDINT(49), "m_udLength",
TO_UDINT(11), "coMerkerEx", TO_UDINT(34), "m_udLength",
TO_UDINT(11), "coRamEx", TO_UDINT(50), "m_udLength",
TO_UDINT(12), "coMerkerEx", TO_UDINT(35), "m_udLength",
TO_UDINT(12), "coRamEx", TO_UDINT(51), "m_udLength",
TO_UDINT(13), "coMerkerEx", TO_UDINT(36), "m_udLength",
TO_UDINT(13), "coRamEx", TO_UDINT(52), "m_udLength",
TO_UDINT(14), "cOnline", TO_UDINT(0), "Online",
TO_UDINT(14), "FwNumStr", TO_UDINT(71), "Data",
TO_UDINT(14), "FwDatetr", TO_UDINT(70), "Data",
TO_UDINT(14), "ToBusIF", TO_UDINT(0), "CallCommand",
TO_UDINT(14), "SdiasIn", TO_UDINT(54), "ClassSvr",
TO_UDINT(15), "cOnline", TO_UDINT(1), "Online",
TO_UDINT(15), "FwNumStr", TO_UDINT(74), "Data",
TO_UDINT(15), "FwDatetr", TO_UDINT(73), "Data",
TO_UDINT(15), "ToBusIF", TO_UDINT(1), "CallCommand",
TO_UDINT(15), "SdiasIn", TO_UDINT(54), "ClassSvr",
TO_UDINT(16), "cOnline", TO_UDINT(2), "Online",
TO_UDINT(16), "FwNumStr", TO_UDINT(77), "Data",
TO_UDINT(16), "FwDatetr", TO_UDINT(76), "Data",
TO_UDINT(16), "ToBusIF", TO_UDINT(2), "CallCommand",
TO_UDINT(16), "SdiasIn", TO_UDINT(54), "ClassSvr",
TO_UDINT(17), "cOnline", TO_UDINT(3), "Online",
TO_UDINT(17), "FwNumStr", TO_UDINT(80), "Data",
TO_UDINT(17), "FwDatetr", TO_UDINT(79), "Data",
TO_UDINT(17), "ToBusIF", TO_UDINT(3), "CallCommand",
TO_UDINT(17), "SdiasIn", TO_UDINT(54), "ClassSvr",
TO_UDINT(21), "To_HwControl", TO_UDINT(26), "Control",
TO_UDINT(24), "SdiasIn", TO_UDINT(54), "ClassSvr",
TO_UDINT(25), "VaranConnect", TO_UDINT(81), "Control",
TO_UDINT(27), "toHwControlBase", TO_UDINT(26), "Control",
TO_UDINT(53), "To_HwControl", TO_UDINT(26), "Control",
TO_UDINT(54), "ToNextSDIAS", TO_UDINT(55), "ClassState",
TO_UDINT(55), "ToBusInterface", TO_UDINT(56), "CallCommand",
TO_UDINT(56), "ToHwControl", TO_UDINT(26), "Control",
TO_UDINT(57), "Current", TO_UDINT(60), "MaxCurrent",
TO_UDINT(58), "SdiasIn", TO_UDINT(54), "ClassSvr",
TO_UDINT(59), "SdiasIn", TO_UDINT(54), "ClassSvr",
TO_UDINT(60), "SdiasIn", TO_UDINT(54), "ClassSvr",
TO_UDINT(61), "SdiasIn", TO_UDINT(54), "ClassSvr",
TO_UDINT(62), "toST151Base", TO_UDINT(60), "ClassState",
TO_UDINT(63), "toST151Base", TO_UDINT(61), "ClassState",
TO_UDINT(64), "DataBuffer", TO_UDINT(28), "m_udLength",
TO_UDINT(65), "DataBuffer", TO_UDINT(29), "m_udLength",
TO_UDINT(66), "DataBuffer", TO_UDINT(30), "m_udLength",
TO_UDINT(67), "DataBuffer", TO_UDINT(31), "m_udLength",
TO_UDINT(68), "DataBuffer", TO_UDINT(32), "m_udLength",
TO_UDINT(69), "DataBuffer", TO_UDINT(37), "m_udLength",
TO_UDINT(70), "DataBuffer", TO_UDINT(38), "m_udLength",
TO_UDINT(71), "DataBuffer", TO_UDINT(39), "m_udLength",
TO_UDINT(72), "DataBuffer", TO_UDINT(40), "m_udLength",
TO_UDINT(73), "DataBuffer", TO_UDINT(41), "m_udLength",
TO_UDINT(74), "DataBuffer", TO_UDINT(42), "m_udLength",
TO_UDINT(75), "DataBuffer", TO_UDINT(43), "m_udLength",
TO_UDINT(76), "DataBuffer", TO_UDINT(44), "m_udLength",
TO_UDINT(77), "DataBuffer", TO_UDINT(45), "m_udLength",
TO_UDINT(78), "DataBuffer", TO_UDINT(46), "m_udLength",
TO_UDINT(79), "DataBuffer", TO_UDINT(47), "m_udLength",
TO_UDINT(80), "DataBuffer", TO_UDINT(48), "m_udLength",
TO_UDINT(81), "To_HwControl", TO_UDINT(26), "Control",

//Initialization values
0$UDINT,
232$UDINT,
TO_UDINT(0), "LEDControl", TO_UDINT(0),//|HW_Network._DriveMng_DC0621\BusInterfaceSdiasDriveMng.LEDControl;
TO_UDINT(0), "Place", TO_UDINT(0),//|HW_Network._DriveMng_DC0621\BusInterfaceSdiasDriveMng.Place;
TO_UDINT(0), "Required", TO_UDINT(1),//|HW_Network._DriveMng_DC0621\BusInterfaceSdiasDriveMng.Required;
TO_UDINT(0), "TimeMultiplier", TO_UDINT(1),//|HW_Network._DriveMng_DC0621\BusInterfaceSdiasDriveMng.TimeMultiplier;
TO_UDINT(0), "SdiasID", TO_UDINT(1801),//|HW_Network._DriveMng_DC0621\BusInterfaceSdiasDriveMng.SdiasID;
TO_UDINT(1), "LEDControl", TO_UDINT(0),//|HW_Network._DriveMng_DC0622\BusInterfaceSdiasDriveMng.LEDControl;
TO_UDINT(1), "Place", TO_UDINT(1),//|HW_Network._DriveMng_DC0622\BusInterfaceSdiasDriveMng.Place;
TO_UDINT(1), "Required", TO_UDINT(1),//|HW_Network._DriveMng_DC0622\BusInterfaceSdiasDriveMng.Required;
TO_UDINT(1), "TimeMultiplier", TO_UDINT(1),//|HW_Network._DriveMng_DC0622\BusInterfaceSdiasDriveMng.TimeMultiplier;
TO_UDINT(1), "SdiasID", TO_UDINT(1801),//|HW_Network._DriveMng_DC0622\BusInterfaceSdiasDriveMng.SdiasID;
TO_UDINT(2), "LEDControl", TO_UDINT(0),//|HW_Network._DriveMng_DC0623\BusInterfaceSdiasDriveMng.LEDControl;
TO_UDINT(2), "Place", TO_UDINT(2),//|HW_Network._DriveMng_DC0623\BusInterfaceSdiasDriveMng.Place;
TO_UDINT(2), "Required", TO_UDINT(1),//|HW_Network._DriveMng_DC0623\BusInterfaceSdiasDriveMng.Required;
TO_UDINT(2), "TimeMultiplier", TO_UDINT(1),//|HW_Network._DriveMng_DC0623\BusInterfaceSdiasDriveMng.TimeMultiplier;
TO_UDINT(2), "SdiasID", TO_UDINT(1801),//|HW_Network._DriveMng_DC0623\BusInterfaceSdiasDriveMng.SdiasID;
TO_UDINT(3), "LEDControl", TO_UDINT(0),//|HW_Network._DriveMng_DC0624\BusInterfaceSdiasDriveMng.LEDControl;
TO_UDINT(3), "Place", TO_UDINT(3),//|HW_Network._DriveMng_DC0624\BusInterfaceSdiasDriveMng.Place;
TO_UDINT(3), "Required", TO_UDINT(1),//|HW_Network._DriveMng_DC0624\BusInterfaceSdiasDriveMng.Required;
TO_UDINT(3), "TimeMultiplier", TO_UDINT(1),//|HW_Network._DriveMng_DC0624\BusInterfaceSdiasDriveMng.TimeMultiplier;
TO_UDINT(3), "SdiasID", TO_UDINT(1801),//|HW_Network._DriveMng_DC0624\BusInterfaceSdiasDriveMng.SdiasID;
TO_UDINT(4), "CanBus", TO_UDINT(0),//|HW_Network._base\CP112_IOs1\_CanLib1.CanBus;
TO_UDINT(5), "CanBus", TO_UDINT(1),//|HW_Network._base\CP112_IOs1\_CanLib2.CanBus;
TO_UDINT(6), "Place", TO_UDINT(0),//|HW_Network._DriveAxis1.Place;
TO_UDINT(6), "AxisNo", TO_UDINT(1),//|HW_Network._DriveAxis1.AxisNo;
TO_UDINT(6), "AxisExtend", TO_UDINT(1),//|HW_Network._DriveAxis1.AxisExtend;
TO_UDINT(6), "ParaSaveType", TO_UDINT(1),//|HW_Network._DriveAxis1.ParaSaveType;
TO_UDINT(6), "OverwriteMotorPara", TO_UDINT(1),//|HW_Network._DriveAxis1.OverwriteMotorPara;
TO_UDINT(7), "Place", TO_UDINT(0),//|HW_Network._DriveAxis2.Place;
TO_UDINT(7), "AxisNo", TO_UDINT(1),//|HW_Network._DriveAxis2.AxisNo;
TO_UDINT(7), "AxisExtend", TO_UDINT(1),//|HW_Network._DriveAxis2.AxisExtend;
TO_UDINT(7), "ParaSaveType", TO_UDINT(1),//|HW_Network._DriveAxis2.ParaSaveType;
TO_UDINT(7), "OverwriteMotorPara", TO_UDINT(1),//|HW_Network._DriveAxis2.OverwriteMotorPara;
TO_UDINT(8), "Place", TO_UDINT(0),//|HW_Network._DriveAxis3.Place;
TO_UDINT(8), "AxisNo", TO_UDINT(1),//|HW_Network._DriveAxis3.AxisNo;
TO_UDINT(8), "AxisExtend", TO_UDINT(1),//|HW_Network._DriveAxis3.AxisExtend;
TO_UDINT(8), "ParaSaveType", TO_UDINT(1),//|HW_Network._DriveAxis3.ParaSaveType;
TO_UDINT(8), "OverwriteMotorPara", TO_UDINT(1),//|HW_Network._DriveAxis3.OverwriteMotorPara;
TO_UDINT(9), "Place", TO_UDINT(0),//|HW_Network._DriveAxis4.Place;
TO_UDINT(9), "AxisNo", TO_UDINT(1),//|HW_Network._DriveAxis4.AxisNo;
TO_UDINT(9), "AxisExtend", TO_UDINT(1),//|HW_Network._DriveAxis4.AxisExtend;
TO_UDINT(9), "ParaSaveType", TO_UDINT(1),//|HW_Network._DriveAxis4.ParaSaveType;
TO_UDINT(9), "OverwriteMotorPara", TO_UDINT(1),//|HW_Network._DriveAxis4.OverwriteMotorPara;
TO_UDINT(10), "ParaSaveType", TO_UDINT(1),//|HW_Network._DriveAxis1\SDDAxSet1.ParaSaveType;
TO_UDINT(10), "OverwriteMotorPara", TO_UDINT(1),//|HW_Network._DriveAxis1\SDDAxSet1.OverwriteMotorPara;
TO_UDINT(11), "ParaSaveType", TO_UDINT(1),//|HW_Network._DriveAxis2\SDDAxSet1.ParaSaveType;
TO_UDINT(11), "OverwriteMotorPara", TO_UDINT(1),//|HW_Network._DriveAxis2\SDDAxSet1.OverwriteMotorPara;
TO_UDINT(12), "ParaSaveType", TO_UDINT(1),//|HW_Network._DriveAxis3\SDDAxSet1.ParaSaveType;
TO_UDINT(12), "OverwriteMotorPara", TO_UDINT(1),//|HW_Network._DriveAxis3\SDDAxSet1.OverwriteMotorPara;
TO_UDINT(13), "ParaSaveType", TO_UDINT(1),//|HW_Network._DriveAxis4\SDDAxSet1.ParaSaveType;
TO_UDINT(13), "OverwriteMotorPara", TO_UDINT(1),//|HW_Network._DriveAxis4\SDDAxSet1.OverwriteMotorPara;
TO_UDINT(14), "Place", TO_UDINT(0),//|HW_Network._DriveMng_DC0621.Place;
TO_UDINT(14), "Required", TO_UDINT(1),//|HW_Network._DriveMng_DC0621.Required;
TO_UDINT(14), "TimeMultiplier", TO_UDINT(1),//|HW_Network._DriveMng_DC0621.TimeMultiplier;
TO_UDINT(15), "Place", TO_UDINT(1),//|HW_Network._DriveMng_DC0622.Place;
TO_UDINT(15), "Required", TO_UDINT(1),//|HW_Network._DriveMng_DC0622.Required;
TO_UDINT(15), "TimeMultiplier", TO_UDINT(1),//|HW_Network._DriveMng_DC0622.TimeMultiplier;
TO_UDINT(16), "Place", TO_UDINT(2),//|HW_Network._DriveMng_DC0623.Place;
TO_UDINT(16), "Required", TO_UDINT(1),//|HW_Network._DriveMng_DC0623.Required;
TO_UDINT(16), "TimeMultiplier", TO_UDINT(1),//|HW_Network._DriveMng_DC0623.TimeMultiplier;
TO_UDINT(17), "Place", TO_UDINT(3),//|HW_Network._DriveMng_DC0624.Place;
TO_UDINT(17), "Required", TO_UDINT(1),//|HW_Network._DriveMng_DC0624.Required;
TO_UDINT(17), "TimeMultiplier", TO_UDINT(1),//|HW_Network._DriveMng_DC0624.TimeMultiplier;
TO_UDINT(18), "Com", TO_UDINT(0),//|HW_Network._base\CP112_IOs1\_SerLib1.Com;
TO_UDINT(19), "Com", TO_UDINT(1),//|HW_Network._base\CP112_IOs1\_SerLib2.Com;
TO_UDINT(24), "LEDControl", TO_UDINT(0),//|HW_Network.DM1611.LEDControl;
TO_UDINT(24), "Place", TO_UDINT(4),//|HW_Network.DM1611.Place;
TO_UDINT(24), "Required", TO_UDINT(1),//|HW_Network.DM1611.Required;
TO_UDINT(25), "Splitter_Place", TO_UDINT(0),//|HW_Network.VaranManager_11\Hub_Base_Root0.Splitter_Place;
TO_UDINT(26), "UdpSafetyPort", TO_UDINT(10823),//|HW_Network.HwControl1.UdpSafetyPort;
TO_UDINT(26), "InterfaceNo", TO_UDINT(1),//|HW_Network.HwControl1.InterfaceNo;
TO_UDINT(28), "ThreadSafe", TO_UDINT(0),//|HW_Network.SerialNoStr\_base\DM1611\MerkerEx0.ThreadSafe;
TO_UDINT(29), "ThreadSafe", TO_UDINT(0),//|HW_Network.SerialNoStr\_base\SR0221\MerkerEx0.ThreadSafe;
TO_UDINT(30), "ThreadSafe", TO_UDINT(0),//|HW_Network.SerialNoStr\_base\ST0111\MerkerEx0.ThreadSafe;
TO_UDINT(31), "ThreadSafe", TO_UDINT(0),//|HW_Network.SerialNoStr\_base\_base\ST1511\MerkerEx0.ThreadSafe;
TO_UDINT(32), "ThreadSafe", TO_UDINT(0),//|HW_Network.SerialNoStr\_base\_base\ST1512\MerkerEx0.ThreadSafe;
TO_UDINT(33), "ThreadSafe", TO_UDINT(0),//|HW_Network._DriveAxis1\MerkerEx2.ThreadSafe;
TO_UDINT(34), "ThreadSafe", TO_UDINT(0),//|HW_Network._DriveAxis2\MerkerEx2.ThreadSafe;
TO_UDINT(35), "ThreadSafe", TO_UDINT(0),//|HW_Network._DriveAxis3\MerkerEx2.ThreadSafe;
TO_UDINT(36), "ThreadSafe", TO_UDINT(0),//|HW_Network._DriveAxis4\MerkerEx2.ThreadSafe;
TO_UDINT(37), "ThreadSafe", TO_UDINT(0),//|HW_Network.SerialNoStr\_base\BusInterfaceSdiasDriveMng\_DriveMng_DC0621\MerkerEx0.ThreadSafe;
TO_UDINT(38), "ThreadSafe", TO_UDINT(0),//|HW_Network.FWDateString\_DriveMng_DC0621\MerkerEx0.ThreadSafe;
TO_UDINT(39), "ThreadSafe", TO_UDINT(0),//|HW_Network.FWNumSTring\_DriveMng_DC0621\MerkerEx0.ThreadSafe;
TO_UDINT(40), "ThreadSafe", TO_UDINT(0),//|HW_Network.SerialNoStr\_base\BusInterfaceSdiasDriveMng\_DriveMng_DC0622\MerkerEx0.ThreadSafe;
TO_UDINT(41), "ThreadSafe", TO_UDINT(0),//|HW_Network.FWDateString\_DriveMng_DC0622\MerkerEx0.ThreadSafe;
TO_UDINT(42), "ThreadSafe", TO_UDINT(0),//|HW_Network.FWNumSTring\_DriveMng_DC0622\MerkerEx0.ThreadSafe;
TO_UDINT(43), "ThreadSafe", TO_UDINT(0),//|HW_Network.SerialNoStr\_base\BusInterfaceSdiasDriveMng\_DriveMng_DC0623\MerkerEx0.ThreadSafe;
TO_UDINT(44), "ThreadSafe", TO_UDINT(0),//|HW_Network.FWDateString\_DriveMng_DC0623\MerkerEx0.ThreadSafe;
TO_UDINT(45), "ThreadSafe", TO_UDINT(0),//|HW_Network.FWNumSTring\_DriveMng_DC0623\MerkerEx0.ThreadSafe;
TO_UDINT(46), "ThreadSafe", TO_UDINT(0),//|HW_Network.SerialNoStr\_base\BusInterfaceSdiasDriveMng\_DriveMng_DC0624\MerkerEx0.ThreadSafe;
TO_UDINT(47), "ThreadSafe", TO_UDINT(0),//|HW_Network.FWDateString\_DriveMng_DC0624\MerkerEx0.ThreadSafe;
TO_UDINT(48), "ThreadSafe", TO_UDINT(0),//|HW_Network.FWNumSTring\_DriveMng_DC0624\MerkerEx0.ThreadSafe;
TO_UDINT(49), "ThreadSafe", TO_UDINT(0),//|HW_Network._DriveAxis1\RAMex2.ThreadSafe;
TO_UDINT(50), "ThreadSafe", TO_UDINT(0),//|HW_Network._DriveAxis2\RAMex2.ThreadSafe;
TO_UDINT(51), "ThreadSafe", TO_UDINT(0),//|HW_Network._DriveAxis3\RAMex2.ThreadSafe;
TO_UDINT(52), "ThreadSafe", TO_UDINT(0),//|HW_Network._DriveAxis4\RAMex2.ThreadSafe;
TO_UDINT(53), "UdpSafetyPort", TO_UDINT(10823),//|HW_Network.HwControl1\SafetyManager.UdpSafetyPort;
TO_UDINT(53), "InterfaceNo", TO_UDINT(1),//|HW_Network.HwControl1\SafetyManager.InterfaceNo;
TO_UDINT(54), "SplitterPlace", TO_UDINT(0),//|HW_Network.SdiasPLC1\SdiasHubBase1.SplitterPlace;
TO_UDINT(55), "DeviceID", TO_UDINT(0),//|HW_Network.SdiasPLC1\SdiasManager1.DeviceID;
TO_UDINT(56), "CycleTime", TO_UDINT(1000),//|HW_Network.SdiasPLC1.CycleTime;
TO_UDINT(56), "IsoStartPoint", TO_UDINT(60),//|HW_Network.SdiasPLC1.IsoStartPoint;
TO_UDINT(58), "LEDControl", TO_UDINT(0),//|HW_Network.SR0221.LEDControl;
TO_UDINT(58), "MinPulse", TO_UDINT(7),//|HW_Network.SR0221.MinPulse;
TO_UDINT(58), "Place", TO_UDINT(6),//|HW_Network.SR0221.Place;
TO_UDINT(58), "Required", TO_UDINT(1),//|HW_Network.SR0221.Required;
TO_UDINT(58), "PWMPeriod", TO_UDINT(32),//|HW_Network.SR0221.PWMPeriod;
TO_UDINT(58), "I2TThreshold", TO_UDINT(100),//|HW_Network.SR0221.I2TThreshold;
TO_UDINT(58), "EncMode", TO_UDINT(1),//|HW_Network.SR0221.EncMode;
TO_UDINT(58), "EncSampling", TO_UDINT(3),//|HW_Network.SR0221.EncSampling;
TO_UDINT(58), "EncDirection", TO_UDINT(0),//|HW_Network.SR0221.EncDirection;
TO_UDINT(58), "InvertZeroPosition", TO_UDINT(0),//|HW_Network.SR0221.InvertZeroPosition;
TO_UDINT(58), "ABCountMode", TO_UDINT(0),//|HW_Network.SR0221.ABCountMode;
TO_UDINT(58), "ExtendedData", TO_UDINT(0),//|HW_Network.SR0221.ExtendedData;
TO_UDINT(59), "LEDControl", TO_UDINT(0),//|HW_Network.ST0111.LEDControl;
TO_UDINT(59), "Place", TO_UDINT(8),//|HW_Network.ST0111.Place;
TO_UDINT(59), "Required", TO_UDINT(1),//|HW_Network.ST0111.Required;
TO_UDINT(59), "UsePulseCntCorrection", TO_UDINT(1),//|HW_Network.ST0111.UsePulseCntCorrection;
TO_UDINT(59), "PulseMode", TO_UDINT(0),//|HW_Network.ST0111.PulseMode;
TO_UDINT(59), "ModeClockCounter", TO_UDINT(0),//|HW_Network.ST0111.ModeClockCounter;
TO_UDINT(59), "InvertEncoder", TO_UDINT(1),//|HW_Network.ST0111.InvertEncoder;
TO_UDINT(59), "InvertEnable", TO_UDINT(1),//|HW_Network.ST0111.InvertEnable;
TO_UDINT(59), "EncoderSampling", TO_UDINT(3),//|HW_Network.ST0111.EncoderSampling;
TO_UDINT(59), "Deathtime", TO_UDINT(60),//|HW_Network.ST0111.Deathtime;
TO_UDINT(59), "Input1Latch", TO_UDINT(0),//|HW_Network.ST0111.Input1Latch;
TO_UDINT(59), "Input2Latch", TO_UDINT(0),//|HW_Network.ST0111.Input2Latch;
TO_UDINT(59), "Input3Latch", TO_UDINT(0),//|HW_Network.ST0111.Input3Latch;
TO_UDINT(59), "ZPulseLatch", TO_UDINT(0),//|HW_Network.ST0111.ZPulseLatch;
TO_UDINT(60), "LEDControl", TO_UDINT(0),//|HW_Network.ST1511.LEDControl;
TO_UDINT(60), "CurrentIncrease", TO_UDINT(1),//|HW_Network.ST1511.CurrentIncrease;
TO_UDINT(60), "HWRampdownDeltaFrequency", TO_UDINT(40),//|HW_Network.ST1511.HWRampdownDeltaFrequency;
TO_UDINT(60), "HWRampdownDeltaTime", TO_UDINT(1),//|HW_Network.ST1511.HWRampdownDeltaTime;
TO_UDINT(60), "CurrentOffsetAdjBridge1", TO_UDINT(100),//|HW_Network.ST1511.CurrentOffsetAdjBridge1;
TO_UDINT(60), "CurrentOffsetAdjBridge2", TO_UDINT(100),//|HW_Network.ST1511.CurrentOffsetAdjBridge2;
TO_UDINT(60), "ChopperOffTime", TO_UDINT(1562),//|HW_Network.ST1511.ChopperOffTime;
TO_UDINT(60), "ChopperOnTimeMin", TO_UDINT(180),//|HW_Network.ST1511.ChopperOnTimeMin;
TO_UDINT(60), "FastDecayTime", TO_UDINT(200),//|HW_Network.ST1511.FastDecayTime;
TO_UDINT(60), "FastDecayTimeFallingStep", TO_UDINT(600),//|HW_Network.ST1511.FastDecayTimeFallingStep;
TO_UDINT(60), "EnableSteps", TO_UDINT(2#1000111),//|HW_Network.ST1511.EnableSteps;
TO_UDINT(60), "FrequLimitIncrease2to1", TO_UDINT(50000),//|HW_Network.ST1511.FrequLimitIncrease2to1;
TO_UDINT(60), "FrequLimitIncrease4to2", TO_UDINT(40000),//|HW_Network.ST1511.FrequLimitIncrease4to2;
TO_UDINT(60), "FrequLimitIncrease8to4", TO_UDINT(30000),//|HW_Network.ST1511.FrequLimitIncrease8to4;
TO_UDINT(60), "FrequLimitIncrease16to8", TO_UDINT(20000),//|HW_Network.ST1511.FrequLimitIncrease16to8;
TO_UDINT(60), "FrequLimitIncrease32to16", TO_UDINT(10000),//|HW_Network.ST1511.FrequLimitIncrease32to16;
TO_UDINT(60), "FrequLimitIncrease64to32", TO_UDINT(5000),//|HW_Network.ST1511.FrequLimitIncrease64to32;
TO_UDINT(60), "FrequLimitDecrease1to2", TO_UDINT(0),//|HW_Network.ST1511.FrequLimitDecrease1to2;
TO_UDINT(60), "FrequLimitDecrease2to4", TO_UDINT(0),//|HW_Network.ST1511.FrequLimitDecrease2to4;
TO_UDINT(60), "FrequLimitDecrease4to8", TO_UDINT(0),//|HW_Network.ST1511.FrequLimitDecrease4to8;
TO_UDINT(60), "FrequLimitDecrease8to16", TO_UDINT(0),//|HW_Network.ST1511.FrequLimitDecrease8to16;
TO_UDINT(60), "FrequLimitDecrease16to32", TO_UDINT(0),//|HW_Network.ST1511.FrequLimitDecrease16to32;
TO_UDINT(60), "FrequLimitDecrease32to64", TO_UDINT(0),//|HW_Network.ST1511.FrequLimitDecrease32to64;
TO_UDINT(60), "Place", TO_UDINT(5),//|HW_Network.ST1511.Place;
TO_UDINT(60), "Required", TO_UDINT(1),//|HW_Network.ST1511.Required;
TO_UDINT(60), "InvertEncoder", TO_UDINT(0),//|HW_Network.ST1511.InvertEncoder;
TO_UDINT(60), "InvertZeroPosition", TO_UDINT(0),//|HW_Network.ST1511.InvertZeroPosition;
TO_UDINT(60), "EncoderSampling", TO_UDINT(3),//|HW_Network.ST1511.EncoderSampling;
TO_UDINT(60), "EncMode", TO_UDINT(0),//|HW_Network.ST1511.EncMode;
TO_UDINT(60), "LatchType", TO_UDINT(0),//|HW_Network.ST1511.LatchType;
TO_UDINT(60), "ABCountMode", TO_UDINT(1),//|HW_Network.ST1511.ABCountMode;
TO_UDINT(60), "StallCurrentReduction", TO_UDINT(0),//|HW_Network.ST1511.StallCurrentReduction;
TO_UDINT(60), "StallCurrentWindow", TO_UDINT(0),//|HW_Network.ST1511.StallCurrentWindow;
TO_UDINT(60), "EnableRegenResistor", TO_UDINT(0),//|HW_Network.ST1511.EnableRegenResistor;
TO_UDINT(60), "RegenResistance", TO_UDINT(150),//|HW_Network.ST1511.RegenResistance;
TO_UDINT(60), "RatedMaxPower", TO_UDINT(1000),//|HW_Network.ST1511.RatedMaxPower;
TO_UDINT(60), "LoadThresholdWarning", TO_UDINT(80),//|HW_Network.ST1511.LoadThresholdWarning;
TO_UDINT(60), "LoadThresholdBridge", TO_UDINT(90),//|HW_Network.ST1511.LoadThresholdBridge;
TO_UDINT(60), "LoadThresholdResistor", TO_UDINT(100),//|HW_Network.ST1511.LoadThresholdResistor;
TO_UDINT(60), "SteppingHysteresis", TO_UDINT(64),//|HW_Network.ST1511.SteppingHysteresis;
TO_UDINT(60), "CompModeVST", TO_UDINT(0),//|HW_Network.ST1511.CompModeVST;
TO_UDINT(60), "UseOszi", TO_UDINT(0),//|HW_Network.ST1511.UseOszi;
TO_UDINT(61), "LEDControl", TO_UDINT(0),//|HW_Network.ST1512.LEDControl;
TO_UDINT(61), "CurrentIncrease", TO_UDINT(1),//|HW_Network.ST1512.CurrentIncrease;
TO_UDINT(61), "HWRampdownDeltaFrequency", TO_UDINT(40),//|HW_Network.ST1512.HWRampdownDeltaFrequency;
TO_UDINT(61), "HWRampdownDeltaTime", TO_UDINT(1),//|HW_Network.ST1512.HWRampdownDeltaTime;
TO_UDINT(61), "CurrentOffsetAdjBridge1", TO_UDINT(100),//|HW_Network.ST1512.CurrentOffsetAdjBridge1;
TO_UDINT(61), "CurrentOffsetAdjBridge2", TO_UDINT(100),//|HW_Network.ST1512.CurrentOffsetAdjBridge2;
TO_UDINT(61), "ChopperOffTime", TO_UDINT(1562),//|HW_Network.ST1512.ChopperOffTime;
TO_UDINT(61), "ChopperOnTimeMin", TO_UDINT(180),//|HW_Network.ST1512.ChopperOnTimeMin;
TO_UDINT(61), "FastDecayTime", TO_UDINT(200),//|HW_Network.ST1512.FastDecayTime;
TO_UDINT(61), "FastDecayTimeFallingStep", TO_UDINT(600),//|HW_Network.ST1512.FastDecayTimeFallingStep;
TO_UDINT(61), "EnableSteps", TO_UDINT(2#1000111),//|HW_Network.ST1512.EnableSteps;
TO_UDINT(61), "FrequLimitIncrease2to1", TO_UDINT(50000),//|HW_Network.ST1512.FrequLimitIncrease2to1;
TO_UDINT(61), "FrequLimitIncrease4to2", TO_UDINT(40000),//|HW_Network.ST1512.FrequLimitIncrease4to2;
TO_UDINT(61), "FrequLimitIncrease8to4", TO_UDINT(30000),//|HW_Network.ST1512.FrequLimitIncrease8to4;
TO_UDINT(61), "FrequLimitIncrease16to8", TO_UDINT(20000),//|HW_Network.ST1512.FrequLimitIncrease16to8;
TO_UDINT(61), "FrequLimitIncrease32to16", TO_UDINT(10000),//|HW_Network.ST1512.FrequLimitIncrease32to16;
TO_UDINT(61), "FrequLimitIncrease64to32", TO_UDINT(5000),//|HW_Network.ST1512.FrequLimitIncrease64to32;
TO_UDINT(61), "FrequLimitDecrease1to2", TO_UDINT(0),//|HW_Network.ST1512.FrequLimitDecrease1to2;
TO_UDINT(61), "FrequLimitDecrease2to4", TO_UDINT(0),//|HW_Network.ST1512.FrequLimitDecrease2to4;
TO_UDINT(61), "FrequLimitDecrease4to8", TO_UDINT(0),//|HW_Network.ST1512.FrequLimitDecrease4to8;
TO_UDINT(61), "FrequLimitDecrease8to16", TO_UDINT(0),//|HW_Network.ST1512.FrequLimitDecrease8to16;
TO_UDINT(61), "FrequLimitDecrease16to32", TO_UDINT(0),//|HW_Network.ST1512.FrequLimitDecrease16to32;
TO_UDINT(61), "FrequLimitDecrease32to64", TO_UDINT(0),//|HW_Network.ST1512.FrequLimitDecrease32to64;
TO_UDINT(61), "Place", TO_UDINT(7),//|HW_Network.ST1512.Place;
TO_UDINT(61), "Required", TO_UDINT(1),//|HW_Network.ST1512.Required;
TO_UDINT(61), "InvertEncoder", TO_UDINT(0),//|HW_Network.ST1512.InvertEncoder;
TO_UDINT(61), "InvertZeroPosition", TO_UDINT(0),//|HW_Network.ST1512.InvertZeroPosition;
TO_UDINT(61), "EncoderSampling", TO_UDINT(3),//|HW_Network.ST1512.EncoderSampling;
TO_UDINT(61), "EncMode", TO_UDINT(0),//|HW_Network.ST1512.EncMode;
TO_UDINT(61), "LatchType", TO_UDINT(0),//|HW_Network.ST1512.LatchType;
TO_UDINT(61), "ABCountMode", TO_UDINT(1),//|HW_Network.ST1512.ABCountMode;
TO_UDINT(61), "StallCurrentReduction", TO_UDINT(0),//|HW_Network.ST1512.StallCurrentReduction;
TO_UDINT(61), "StallCurrentWindow", TO_UDINT(0),//|HW_Network.ST1512.StallCurrentWindow;
TO_UDINT(61), "EnableRegenResistor", TO_UDINT(0),//|HW_Network.ST1512.EnableRegenResistor;
TO_UDINT(61), "RegenResistance", TO_UDINT(150),//|HW_Network.ST1512.RegenResistance;
TO_UDINT(61), "RatedMaxPower", TO_UDINT(1000),//|HW_Network.ST1512.RatedMaxPower;
TO_UDINT(61), "LoadThresholdWarning", TO_UDINT(80),//|HW_Network.ST1512.LoadThresholdWarning;
TO_UDINT(61), "LoadThresholdBridge", TO_UDINT(90),//|HW_Network.ST1512.LoadThresholdBridge;
TO_UDINT(61), "LoadThresholdResistor", TO_UDINT(100),//|HW_Network.ST1512.LoadThresholdResistor;
TO_UDINT(61), "SteppingHysteresis", TO_UDINT(64),//|HW_Network.ST1512.SteppingHysteresis;
TO_UDINT(61), "CompModeVST", TO_UDINT(0),//|HW_Network.ST1512.CompModeVST;
TO_UDINT(61), "UseOszi", TO_UDINT(0),//|HW_Network.ST1512.UseOszi;
TO_UDINT(64), "SingleRealloc", TO_UDINT(1),//|HW_Network._base\DM1611\SerialNoStr.SingleRealloc;
TO_UDINT(65), "SingleRealloc", TO_UDINT(1),//|HW_Network._base\SR0221\SerialNoStr.SingleRealloc;
TO_UDINT(66), "SingleRealloc", TO_UDINT(1),//|HW_Network._base\ST0111\SerialNoStr.SingleRealloc;
TO_UDINT(67), "SingleRealloc", TO_UDINT(1),//|HW_Network._base\_base\ST1511\SerialNoStr.SingleRealloc;
TO_UDINT(68), "SingleRealloc", TO_UDINT(1),//|HW_Network._base\_base\ST1512\SerialNoStr.SingleRealloc;
TO_UDINT(69), "SingleRealloc", TO_UDINT(1),//|HW_Network._base\BusInterfaceSdiasDriveMng\_DriveMng_DC0621\SerialNoStr.SingleRealloc;
TO_UDINT(70), "SingleRealloc", TO_UDINT(1),//|HW_Network._DriveMng_DC0621\FWDateString.SingleRealloc;
TO_UDINT(71), "SingleRealloc", TO_UDINT(1),//|HW_Network._DriveMng_DC0621\FWNumSTring.SingleRealloc;
TO_UDINT(72), "SingleRealloc", TO_UDINT(1),//|HW_Network._base\BusInterfaceSdiasDriveMng\_DriveMng_DC0622\SerialNoStr.SingleRealloc;
TO_UDINT(73), "SingleRealloc", TO_UDINT(1),//|HW_Network._DriveMng_DC0622\FWDateString.SingleRealloc;
TO_UDINT(74), "SingleRealloc", TO_UDINT(1),//|HW_Network._DriveMng_DC0622\FWNumSTring.SingleRealloc;
TO_UDINT(75), "SingleRealloc", TO_UDINT(1),//|HW_Network._base\BusInterfaceSdiasDriveMng\_DriveMng_DC0623\SerialNoStr.SingleRealloc;
TO_UDINT(76), "SingleRealloc", TO_UDINT(1),//|HW_Network._DriveMng_DC0623\FWDateString.SingleRealloc;
TO_UDINT(77), "SingleRealloc", TO_UDINT(1),//|HW_Network._DriveMng_DC0623\FWNumSTring.SingleRealloc;
TO_UDINT(78), "SingleRealloc", TO_UDINT(1),//|HW_Network._base\BusInterfaceSdiasDriveMng\_DriveMng_DC0624\SerialNoStr.SingleRealloc;
TO_UDINT(79), "SingleRealloc", TO_UDINT(1),//|HW_Network._DriveMng_DC0624\FWDateString.SingleRealloc;
TO_UDINT(80), "SingleRealloc", TO_UDINT(1),//|HW_Network._DriveMng_DC0624\FWNumSTring.SingleRealloc;
TO_UDINT(81), "VaranManagerTime", TO_UDINT(1000000),//|HW_Network.VaranManager_11.VaranManagerTime;
TO_UDINT(81), "VaranManagerNr", TO_UDINT(0),//|HW_Network.VaranManager_11.VaranManagerNr;
TO_UDINT(81), "PayloadFrame", TO_UDINT(0),//|HW_Network.VaranManager_11.PayloadFrame;
TO_UDINT(81), "CoreSelect", TO_UDINT(0),//|HW_Network.VaranManager_11.CoreSelect;

//Symbolic initialization values
0$UDINT,
0$UDINT,

//Initialization of string values
0$UDINT,
0$UDINT,

//Configuration of tasks (RealTime, Cyclic, Background)
0$UDINT,
1$UDINT,
TO_UDINT(27), (1)$UDINT, 4194304$DINT, 	//HWCONTROL1\HWRTPOSTSCAN

0$UDINT,
4$UDINT,
TO_UDINT(14), (10)$UDINT, 4194303$DINT, 	//_DRIVEMNG_DC0621
TO_UDINT(15), (10)$UDINT, 4194303$DINT, 	//_DRIVEMNG_DC0622
TO_UDINT(16), (10)$UDINT, 4194303$DINT, 	//_DRIVEMNG_DC0623
TO_UDINT(17), (10)$UDINT, 4194303$DINT, 	//_DRIVEMNG_DC0624

0$UDINT,
0$UDINT,

//External connections
0$UDINT,
0$UDINT,

//Magic internal connections
0$UDINT,
39$UDINT,
TO_UDINT(0), "SdiasIn", TO_UDINT(14), "SdiasIn",
TO_UDINT(0), "Place", TO_UDINT(14), "Place",
TO_UDINT(0), "Required", TO_UDINT(14), "Required",
TO_UDINT(0), "TimeMultiplier", TO_UDINT(14), "TimeMultiplier",
TO_UDINT(1), "SdiasIn", TO_UDINT(15), "SdiasIn",
TO_UDINT(1), "Place", TO_UDINT(15), "Place",
TO_UDINT(1), "Required", TO_UDINT(15), "Required",
TO_UDINT(1), "TimeMultiplier", TO_UDINT(15), "TimeMultiplier",
TO_UDINT(2), "SdiasIn", TO_UDINT(16), "SdiasIn",
TO_UDINT(2), "Place", TO_UDINT(16), "Place",
TO_UDINT(2), "Required", TO_UDINT(16), "Required",
TO_UDINT(2), "TimeMultiplier", TO_UDINT(16), "TimeMultiplier",
TO_UDINT(3), "SdiasIn", TO_UDINT(17), "SdiasIn",
TO_UDINT(3), "Place", TO_UDINT(17), "Place",
TO_UDINT(3), "Required", TO_UDINT(17), "Required",
TO_UDINT(3), "TimeMultiplier", TO_UDINT(17), "TimeMultiplier",
TO_UDINT(10), "ParaSaveType", TO_UDINT(6), "ParaSaveType",
TO_UDINT(10), "OverwriteMotorPara", TO_UDINT(6), "OverwriteMotorPara",
TO_UDINT(10), "ParaTab", TO_UDINT(6), "ParaTab",
TO_UDINT(10), "FileHandle", TO_UDINT(6), "FileHandle",
TO_UDINT(10), "TableIndex", TO_UDINT(6), "TableIndex",
TO_UDINT(11), "ParaSaveType", TO_UDINT(7), "ParaSaveType",
TO_UDINT(11), "OverwriteMotorPara", TO_UDINT(7), "OverwriteMotorPara",
TO_UDINT(11), "ParaTab", TO_UDINT(7), "ParaTab",
TO_UDINT(11), "FileHandle", TO_UDINT(7), "FileHandle",
TO_UDINT(11), "TableIndex", TO_UDINT(7), "TableIndex",
TO_UDINT(12), "ParaSaveType", TO_UDINT(8), "ParaSaveType",
TO_UDINT(12), "OverwriteMotorPara", TO_UDINT(8), "OverwriteMotorPara",
TO_UDINT(12), "ParaTab", TO_UDINT(8), "ParaTab",
TO_UDINT(12), "FileHandle", TO_UDINT(8), "FileHandle",
TO_UDINT(12), "TableIndex", TO_UDINT(8), "TableIndex",
TO_UDINT(13), "ParaSaveType", TO_UDINT(9), "ParaSaveType",
TO_UDINT(13), "OverwriteMotorPara", TO_UDINT(9), "OverwriteMotorPara",
TO_UDINT(13), "ParaTab", TO_UDINT(9), "ParaTab",
TO_UDINT(13), "FileHandle", TO_UDINT(9), "FileHandle",
TO_UDINT(13), "TableIndex", TO_UDINT(9), "TableIndex",
TO_UDINT(53), "UdpSafetyPort", TO_UDINT(26), "UdpSafetyPort",
TO_UDINT(53), "InterfaceNo", TO_UDINT(26), "InterfaceNo",
TO_UDINT(53), "SafetyDomainTimeout", TO_UDINT(26), "SafetyDomainTimeout",

//Configuration of timeslots of tasks (RealTime, Cyclic)
#ifdef __LSLLDR_TIMESLOTS__
0$UDINT,
0$UDINT,

0$UDINT,
0$UDINT,

#endif //__LSLLDR_TIMESLOTS__

//MultiMaster connections
#ifdef __LSLLDR_MULTIMASTER__
0$UDINT,
0$UDINT,
#endif //__LSLLDR_MULTIMASTER__

//Configuration for task ID (RealTime, CyclicTime)
#ifdef __LSLLDR_TASKID__
"\\\\TASKS2  "
0$UDINT,
1$UDINT,
(0)$UDINT, 	//HWCONTROL1\HWRTPOSTSCAN

0$UDINT,
4$UDINT,
(0)$UDINT, 	//_DRIVEMNG_DC0621
(0)$UDINT, 	//_DRIVEMNG_DC0622
(0)$UDINT, 	//_DRIVEMNG_DC0623
(0)$UDINT, 	//_DRIVEMNG_DC0624

0$UDINT,
0$UDINT,

#endif //__LSLLDR_TASKID__

END_FUNCTION
